(* IEC 61131-3 sources: llm-plc-st-eval/data/definitivo/claude-sonnet-4-6/B5/zero_shot, 3 files *)

(* ---- ejec_1.st ---- *)
```pascal
FUNCTION_BLOCK FB_Ventilador
VAR_INPUT
    quemadorOn : BOOL; (* Señal del quemador: TRUE = encendido *)
END_VAR

VAR_OUTPUT
    ventilador : BOOL; (* Salida del ventilador: TRUE = funcionando *)
END_VAR

VAR
    tonApagado : TON;  (* Temporizador de retardo al apagado *)
END_VAR

(*
    Lógica:
    - Si el quemador está encendido, el ventilador funciona y el temporizador se mantiene reseteado.
    - Al apagarse el quemador, el temporizador inicia el conteo de 30 s.
    - Cuando el temporizador completa los 30 s (Q = TRUE), el ventilador se detiene.
*)

(* Activar temporizador solo cuando el quemador está apagado *)
tonApagado(
    IN := NOT quemadorOn,
    PT := T#30S
);

(* El ventilador funciona si el quemador está encendido
   O si el temporizador aún no ha completado los 30 s *)
ventilador := quemadorOn OR (NOT tonApagado.Q);

END_FUNCTION_BLOCK
```

(* ---- ejec_2.st ---- *)
```pascal
FUNCTION_BLOCK FB_Ventilador
VAR_INPUT
    quemadorOn : BOOL; (* Señal del quemador: TRUE = encendido *)
END_VAR

VAR_OUTPUT
    ventilador : BOOL; (* Salida del ventilador: TRUE = funcionando *)
END_VAR

VAR
    tonPostApagado : TON;  (* Temporizador de retardo al apagado *)
END_VAR

(* -------------------------------------------------------
   Lógica:
   - Quemador ON  → ventilador ON, temporizador en reset.
   - Quemador OFF → temporizador inicia 30 s; ventilador
     permanece ON hasta que el temporizador expire.
   ------------------------------------------------------- *)

(* Activar temporizador solo cuando el quemador está apagado *)
tonPostApagado(
    IN  := NOT quemadorOn,  (* Cuenta mientras quemador esté OFF *)
    PT  := T#30S            (* Tiempo de post-ventilación *)
);

(* El ventilador funciona si el quemador está ON
   o si el temporizador aún no ha expirado *)
ventilador := quemadorOn OR NOT tonPostApagado.Q;

END_FUNCTION_BLOCK
```

(* ---- ejec_3.st ---- *)
```pascal
FUNCTION_BLOCK FB_Ventilador
VAR_INPUT
    quemadorOn : BOOL; (* Señal del quemador: TRUE = encendido *)
END_VAR

VAR_OUTPUT
    ventilador : BOOL; (* Salida del ventilador: TRUE = funcionando *)
END_VAR

VAR
    tonPostApagado : TON;  (* Temporizador de retardo al apagado *)
END_VAR

(*
    Lógica:
    - Si el quemador está encendido, el ventilador funciona y el temporizador se mantiene reseteado.
    - Al apagarse el quemador, el temporizador comienza a contar 30 segundos.
    - Cuando el temporizador completa los 30 segundos (Q = TRUE), el ventilador se detiene.
*)

(* Activar temporizador solo cuando el quemador está apagado *)
tonPostApagado(
    IN  := NOT quemadorOn,  (* Inicia cuenta cuando el quemador se apaga *)
    PT  := T#30S            (* Tiempo de post-ventilación: 30 segundos   *)
);

(* El ventilador funciona si el quemador está ON,
   o si el temporizador aún no ha completado los 30 s *)
ventilador := quemadorOn OR NOT tonPostApagado.Q;
```
